(* IEC 61131-3 sources: plc-iiot-stack/src/POUs/Json/F_IsFiniteLreal, 1 file *)

(* ---- F_IsFiniteLreal.decl.st ---- *)
// Назначение: проверка, что LREAL — конечное число (не NaN и не бесконечность): порядок не из одних единиц.
// Автор:      kr0nsch
// Версия:     0.1.0
// Документ:   docs/plc_mqtt.md, раздел «Построение JSON»
FUNCTION F_IsFiniteLreal : BOOL
VAR_INPUT
    lrValue : LREAL;
END_VAR
VAR
    pBits : POINTER TO LWORD;   // те же 8 байт, что lrValue
END_VAR
